// Optional read-only status of a telescope control, for the HMI gateway (why not ready, last rejected command, current
// position). Separate from the I_Telescope hierarchy on purpose: it does not extend I_Telescope, so an implementation that
// does not provide it is not forced to. specs/design/ui-tiers-and-hmi-gateway.md, section 3.1.
INTERFACE I_TelescopeStatus

// A component of the telescope is in error.
PROPERTY Error : BOOL
GET
END_GET
END_PROPERTY

// Error number of that component.
PROPERTY ErrorID : UDINT
GET
END_GET
END_PROPERTY

// A command sequence is running (power-on, park, slew, goto, home, stop).
PROPERTY Busy : BOOL
GET
END_GET
END_PROPERTY

// The telescope is parked.
PROPERTY IsParked : BOOL
GET
END_GET
END_PROPERTY

// The telescope state machine does not run (MONET manual mode).
PROPERTY Suspended : BOOL
GET
END_GET
END_PROPERTY

// The command the telescope refused last.
PROPERTY LastRejectedCommand : E_TCSCommand
GET
END_GET
END_PROPERTY

// Why it refused it (F_CommandAcceptance).
PROPERTY LastRejectReason : E_CommandRejectReason
GET
END_GET
END_PROPERTY

// +1 per rejected command; a consumer detects a new rejection by the change.
PROPERTY RejectCount : UDINT
GET
END_GET
END_PROPERTY

// deg, ICRS, current position of the axes (not the target).
PROPERTY CurrentRightAscension : LREAL
GET
END_GET
END_PROPERTY

// deg, ICRS, current position of the axes (not the target).
PROPERTY CurrentDeclination : LREAL
GET
END_GET
END_PROPERTY

END_INTERFACE

(* stored: Version 1.1.0.1, ProductVersion 3.1.4024.15
   Itf I_TelescopeStatus: Id {e7f9a0ad-cbab-4b11-8040-faf0a9882628}
   Property Error: Id {21845583-423b-44b3-9517-82fb2eba08ec}
   Get Get: Id {0ea8eda4-f9c8-4302-b77e-71d643e5c992}
   Property ErrorID: Id {2f8af68d-784d-422c-95cc-78131eca57fc}
   Get Get: Id {8dab492c-a457-4dbd-aa5b-50bd510cc880}
   Property Busy: Id {2b5c42a4-6376-45de-93bf-2b470a57603c}
   Get Get: Id {2e58cf32-ba06-4c4b-801d-0acc4e0fc5e9}
   Property IsParked: Id {1e5508de-10dc-4883-b5d8-5097131380cc}
   Get Get: Id {327d1f4c-2175-4e84-bc0d-fea2eeed5c3d}
   Property Suspended: Id {d22ab7f4-a5d2-4c5e-8679-c71af16710cd}
   Get Get: Id {588a541f-bf94-46f3-8e29-5042a25edc7b}
   Property LastRejectedCommand: Id {fe0da4e3-846d-43dc-8a67-d682e3ab8252}
   Get Get: Id {550ebfee-b371-4c40-acf6-4e460e71e605}
   Property LastRejectReason: Id {65c7239d-e495-4455-94b1-824a24fcce98}
   Get Get: Id {91d0af8c-dc2f-497a-b594-19543cec9b0b}
   Property RejectCount: Id {2a4c511c-4fca-4b80-800d-7804b68798f2}
   Get Get: Id {a1f3f7e4-07c8-44fa-a899-e4549e8c2fa1}
   Property CurrentRightAscension: Id {8d37c925-14c9-4a6f-bae5-576e82e5bd7d}
   Get Get: Id {293fceec-932a-4a54-aec0-e9f6ae789c26}
   Property CurrentDeclination: Id {bfef482b-165b-4056-a3a6-04624ff32c20}
   Get Get: Id {d6b937a3-b242-438a-b4ea-efe6f5099d35} *)
